(* PLC project fwd_rev_interlock, Unknown Lessons in Electric Circuits transcription 1 *)
(* stored: creationDateTime 2026-09-02T12:00:00 *)

PROGRAM main
  VAR
    START_FWD : BOOL;
    START_REV : BOOL;
    STOP : BOOL;
    M1_FWD : BOOL;
    M2_REV : BOOL;
  END_VAR

(* LD diagram, written out as Structured Text *)
M1_FWD := (START_FWD OR M1_FWD) AND NOT STOP AND NOT M2_REV;
M2_REV := (START_REV OR M2_REV) AND NOT STOP AND NOT M1_FWD;
END_PROGRAM

CONFIGURATION Config0
  RESOURCE Res0 ON PLC
    TASK tcyclic(INTERVAL := T#10ms, PRIORITY := 0);
    PROGRAM inst0 WITH tcyclic : main;
  END_RESOURCE
END_CONFIGURATION
